// TIA Portal V20 export
// export: Created 2026-10-19T18:06:21.5238281Z, ExportSetting WithDefaults, DisplayName Totally Integrated Automation Portal, DisplayVersion V20 Update 6, DisplayName TIA Portal Openness, DisplayVersion V20 Update 6, DisplayName TIA Portal Version Control Interface, DisplayVersion V20 Update 6, DisplayName SINAMICS Startdrive Advanced, DisplayVersion V20 SP1, DisplayName SINAMICS Startdrive G130, G150, S120, S150, SINAMICS MV, G220, S200, S210, DisplayVersion V20 SP1, DisplayName SINAMICS Startdrive G110M, G120, G120C, G120D, G120P, G115D, DisplayVersion V20 SP1, DisplayName STEP 7 Professional, DisplayVersion V20 Update 6, DisplayName STEP 7 Safety, DisplayVersion V20 Update 2, DisplayName WinCC Basic/Comfort/Advanced, DisplayVersion V20 Update 6, DisplayName WinCC Unified, DisplayVersion V20 Update 6
FUNCTION_BLOCK "SAI_IND_CalFree"   // FB53, LAD
TITLE = CalFree Adjustment
{ S7_Optimized_Access := 'FALSE' }
VERSION : 0.1
// CalFree is a method of analog scale adjustment without using test weights. It takes the factory calibrated load cell Rated Output (mV/ Vexc.) and user defined scale capacity to build a linear loading curve.
// This method is usually applied to huge capacity scales in which calibration with test weights or other material is not feasible at all.
// stored: AutoNumber true, IsIECCheckEnabled false, SetENOAutomatically false, UDAEnableTagReadback false
   VAR_INPUT
      ID : HW_IO;   // The Profinet Device Hardware Identifier under device properties
   END_VAR
   VAR_OUTPUT
      Process : Bool;   // Adjustment is in process
      Done : Bool;   // Adjustment completed successfully
      Error : Bool;
   END_VAR
   VAR_IN_OUT
      RatedCapacity : Real;   // Scale Capacity
      Unit : SInt := 1;   // Decimal 0 - gram; 1 - KG; 2 - Lbs
      RatedOutput : Real;   // The averaged load cells' Rated Output in mV/V
      Start : Bool;   // Switch ON to start adjustment
   END_VAR
   VAR DB_SPECIFIC
      Activate : Bool;
      Status_RECORD : Int;
      CalFree_RECORD : Int;
      AdjustStep : SInt;
      Check01 : Bool;
      Check02 : Bool;
   END_VAR
   VAR
      WRREC_CalFree { S7_SetPoint := 'True'} : WRREC;
   END_VAR
   VAR DB_SPECIFIC
      Static01 : Bool;
   END_VAR
   VAR
      RDREC_Status { S7_SetPoint := 'True'} : RDREC;
   END_VAR
   VAR_TEMP   // added for the SCL form of the ladder/FBD networks
      _w1 : Bool;
      _w2 : Bool;
      _w3 : Bool;
      _w4 : Bool;
      _w5 : Bool;
      _w6 : Bool;
      _w7 : Bool;
      _w8 : Bool;
      _w9 : Bool;
      _w10 : Bool;
      _w11 : Bool;
   END_VAR
BEGIN

REGION Network 1: Start routine
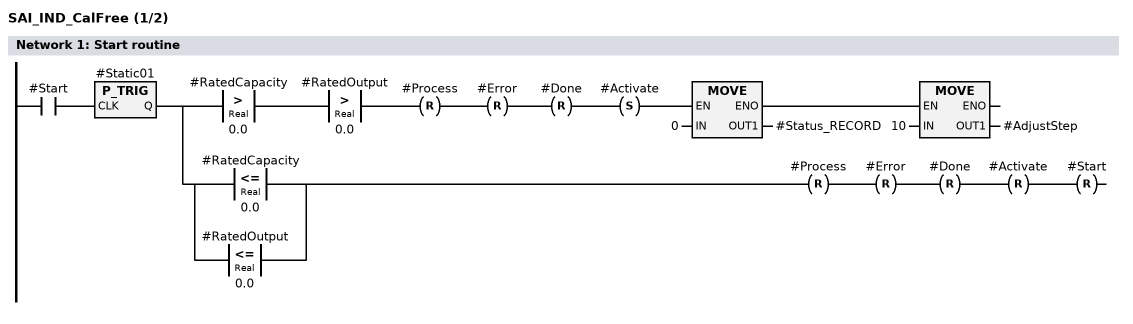
   RUNG wire#powerrail
      Contact( #Start )
      P_Trig( #Static01 )
      wire#w1
      { S7_Templates := "SrcType := Real" } GT_Contact(in1 := #RatedCapacity, in2 := 0.0)
      { S7_Templates := "SrcType := Real" } GT_Contact(in1 := #RatedOutput, in2 := 0.0)
      R_Coil( #Process )
      R_Coil( #Error )
      R_Coil( #Done )
      S_Coil( #Activate )
      Move(in := 0, out1 => #Status_RECORD)
      Move(in := 10, out1 => #AdjustStep)
   END_RUNG
   RUNG wire#w1
      { S7_Templates := "SrcType := Real" } LE_Contact(in1 := #RatedCapacity, in2 := 0.0)
      wire#w2
      R_Coil( #Process )
      R_Coil( #Error )
      R_Coil( #Done )
      R_Coil( #Activate )
      R_Coil( #Start )
   END_RUNG
   RUNG wire#w1
      { S7_Templates := "SrcType := Real" } LE_Contact(in1 := #RatedOutput, in2 := 0.0)
   END_RUNG wire#w2
   // the same network as SCL:
   #_w1 := #Start AND NOT #Static01;   // rising edge
   #Static01 := #Start;
   IF #_w1 AND (#RatedCapacity > 0.0) AND (#RatedOutput > 0.0) THEN
       #Process := FALSE;
       #Error := FALSE;
       #Done := FALSE;
       #Activate := TRUE;
       #Status_RECORD := 0;
       #AdjustStep := 10;
   END_IF;
   IF #_w1 AND ((#RatedCapacity <= 0.0) OR (#RatedOutput <= 0.0)) THEN
       #Process := FALSE;
       #Error := FALSE;
       #Done := FALSE;
       #Activate := FALSE;
       #Start := FALSE;
   END_IF;
END_REGION

REGION Network 2: Sequence
   // CalFree adjustment steps:
   // 
   // 1. Switch on Input bit Start
   // 
   // 2. Write in (a) Scale Capacity (Index 0x401A), (b) Scale unit (Index 0x401C, Decimal 0 - gram; Decimal 1 - KG; Decimal 2 - Pounds) and (c) Load Cells' averaged Rated Output (Index 0x401D, in mV/V)
   // 
   // 3. Start CalFree adjustment (Index 0x401A)
   // 
   // 4. Continuously read in adjustment status (Index 0x4007)
   // 
   // 5. Output bit Done will be turned ON after completion of the process
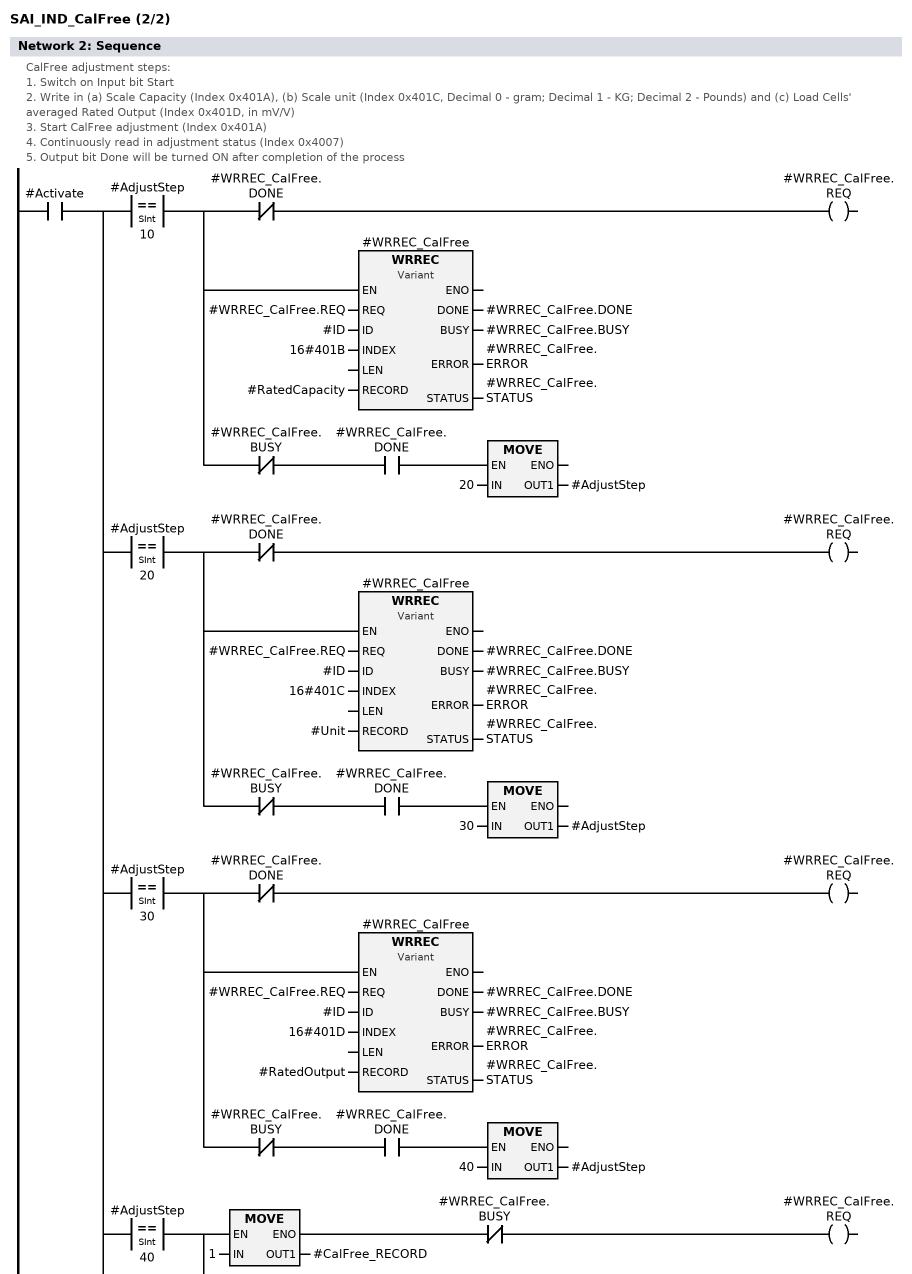
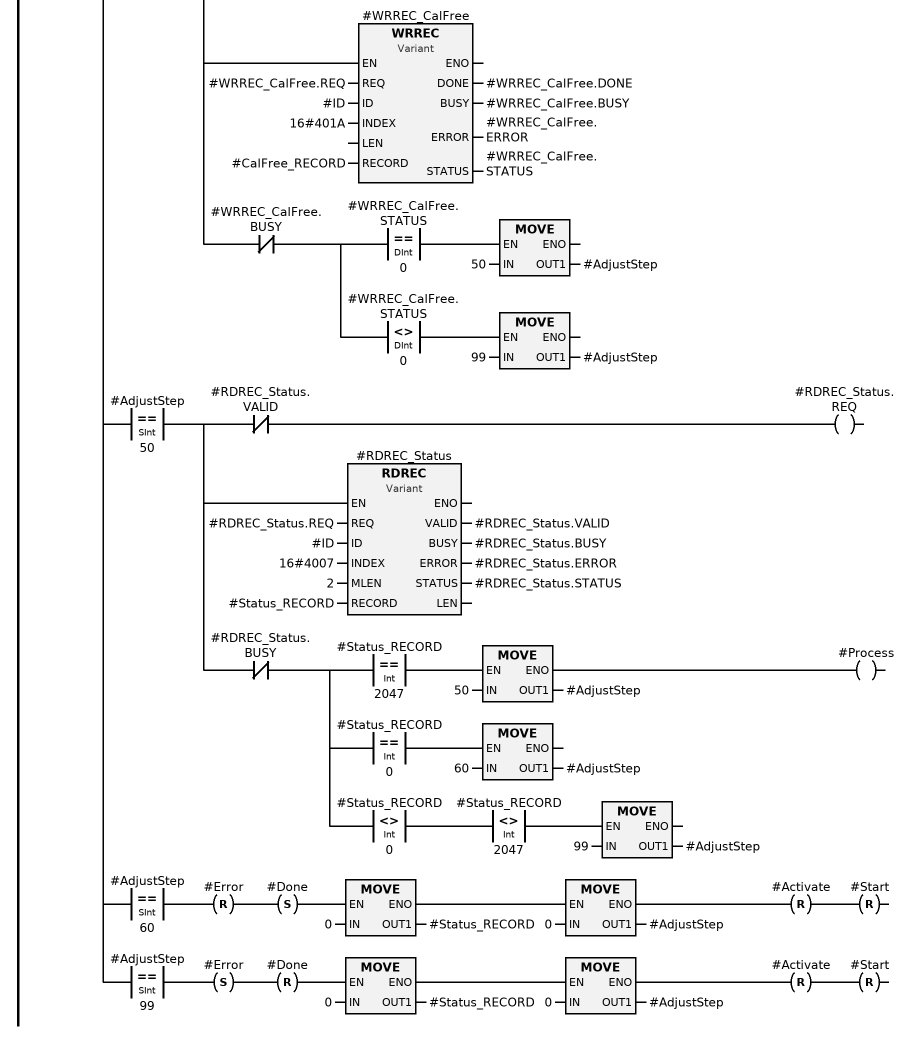
   RUNG wire#powerrail
      Contact( #Activate )
      wire#w1
      { S7_Templates := "SrcType := SInt" } EQ_Contact(in1 := #AdjustStep, in2 := 10)
      wire#w2
      I_Contact( #WRREC_CalFree.DONE )
      Coil( #WRREC_CalFree.REQ )
   END_RUNG
   RUNG wire#w2
      { S7_Templates := "[ptr_type := Variant, id_type := HW_IO, index_type := DInt, len_type := UInt]" } #WRREC_CalFree.WRREC(REQ := #WRREC_CalFree.REQ, ID := #ID, INDEX := 16#401B, LEN :=, RECORD := #RatedCapacity, DONE => #WRREC_CalFree.DONE, BUSY => #WRREC_CalFree.BUSY, ERROR => #WRREC_CalFree.ERROR, STATUS => #WRREC_CalFree.STATUS)
   END_RUNG
   RUNG wire#w2
      I_Contact( #WRREC_CalFree.BUSY )
      Contact( #WRREC_CalFree.DONE )
      Move(in := 20, out1 => #AdjustStep)
   END_RUNG
   RUNG wire#w1
      { S7_Templates := "SrcType := SInt" } EQ_Contact(in1 := #AdjustStep, in2 := 20)
      wire#w3
      I_Contact( #WRREC_CalFree.DONE )
      Coil( #WRREC_CalFree.REQ )
   END_RUNG
   RUNG wire#w3
      { S7_Templates := "[ptr_type := Variant, id_type := HW_IO, index_type := DInt, len_type := UInt]" } #WRREC_CalFree.WRREC(REQ := #WRREC_CalFree.REQ, ID := #ID, INDEX := 16#401C, LEN :=, RECORD := #Unit, DONE => #WRREC_CalFree.DONE, BUSY => #WRREC_CalFree.BUSY, ERROR => #WRREC_CalFree.ERROR, STATUS => #WRREC_CalFree.STATUS)
   END_RUNG
   RUNG wire#w3
      I_Contact( #WRREC_CalFree.BUSY )
      Contact( #WRREC_CalFree.DONE )
      Move(in := 30, out1 => #AdjustStep)
   END_RUNG
   RUNG wire#w1
      { S7_Templates := "SrcType := SInt" } EQ_Contact(in1 := #AdjustStep, in2 := 30)
      wire#w4
      I_Contact( #WRREC_CalFree.DONE )
      Coil( #WRREC_CalFree.REQ )
   END_RUNG
   RUNG wire#w4
      { S7_Templates := "[ptr_type := Variant, id_type := HW_IO, index_type := DInt, len_type := UInt]" } #WRREC_CalFree.WRREC(REQ := #WRREC_CalFree.REQ, ID := #ID, INDEX := 16#401D, LEN :=, RECORD := #RatedOutput, DONE => #WRREC_CalFree.DONE, BUSY => #WRREC_CalFree.BUSY, ERROR => #WRREC_CalFree.ERROR, STATUS => #WRREC_CalFree.STATUS)
   END_RUNG
   RUNG wire#w4
      I_Contact( #WRREC_CalFree.BUSY )
      Contact( #WRREC_CalFree.DONE )
      Move(in := 40, out1 => #AdjustStep)
   END_RUNG
   RUNG wire#w1
      { S7_Templates := "SrcType := SInt" } EQ_Contact(in1 := #AdjustStep, in2 := 40)
      wire#w5
      Move(in := 1, out1 => #CalFree_RECORD)
      I_Contact( #WRREC_CalFree.BUSY )
      Coil( #WRREC_CalFree.REQ )
   END_RUNG
   RUNG wire#w5
      { S7_Templates := "[ptr_type := Variant, id_type := HW_IO, index_type := DInt, len_type := UInt]" } #WRREC_CalFree.WRREC(REQ := #WRREC_CalFree.REQ, ID := #ID, INDEX := 16#401A, LEN :=, RECORD := #CalFree_RECORD, DONE => #WRREC_CalFree.DONE, BUSY => #WRREC_CalFree.BUSY, ERROR => #WRREC_CalFree.ERROR, STATUS => #WRREC_CalFree.STATUS)
   END_RUNG
   RUNG wire#w5
      I_Contact( #WRREC_CalFree.BUSY )
      wire#w6
      { S7_Templates := "SrcType := DInt" } EQ_Contact(in1 := #WRREC_CalFree.STATUS, in2 := 0)
      Move(in := 50, out1 => #AdjustStep)
   END_RUNG
   RUNG wire#w6
      { S7_Templates := "SrcType := DInt" } NE_Contact(in1 := #WRREC_CalFree.STATUS, in2 := 0)
      Move(in := 99, out1 => #AdjustStep)
   END_RUNG
   RUNG wire#w1
      { S7_Templates := "SrcType := SInt" } EQ_Contact(in1 := #AdjustStep, in2 := 50)
      wire#w7
      I_Contact( #RDREC_Status.VALID )
      Coil( #RDREC_Status.REQ )
   END_RUNG
   RUNG wire#w7
      { S7_Templates := "[ptr_type := Variant, id_type := HW_IO, index_type := DInt, len_type := UInt]" } #RDREC_Status.RDREC(REQ := #RDREC_Status.REQ, ID := #ID, INDEX := 16#4007, MLEN := 2, RECORD := #Status_RECORD, VALID => #RDREC_Status.VALID, BUSY => #RDREC_Status.BUSY, ERROR => #RDREC_Status.ERROR, STATUS => #RDREC_Status.STATUS, LEN =>)
   END_RUNG
   RUNG wire#w7
      I_Contact( #RDREC_Status.BUSY )
      wire#w8
      { S7_Templates := "SrcType := Int" } EQ_Contact(in1 := #Status_RECORD, in2 := 2047)
      Move(in := 50, out1 => #AdjustStep)
      Coil( #Process )
   END_RUNG
   RUNG wire#w8
      { S7_Templates := "SrcType := Int" } EQ_Contact(in1 := #Status_RECORD, in2 := 0)
      Move(in := 60, out1 => #AdjustStep)
   END_RUNG
   RUNG wire#w8
      { S7_Templates := "SrcType := Int" } NE_Contact(in1 := #Status_RECORD, in2 := 0)
      { S7_Templates := "SrcType := Int" } NE_Contact(in1 := #Status_RECORD, in2 := 2047)
      Move(in := 99, out1 => #AdjustStep)
   END_RUNG
   RUNG wire#w1
      { S7_Templates := "SrcType := SInt" } EQ_Contact(in1 := #AdjustStep, in2 := 60)
      R_Coil( #Error )
      S_Coil( #Done )
      Move(in := 0, out1 => #Status_RECORD)
      Move(in := 0, out1 => #AdjustStep)
      R_Coil( #Activate )
      R_Coil( #Start )
   END_RUNG
   RUNG wire#w1
      { S7_Templates := "SrcType := SInt" } EQ_Contact(in1 := #AdjustStep, in2 := 99)
      S_Coil( #Error )
      R_Coil( #Done )
      Move(in := 0, out1 => #Status_RECORD)
      Move(in := 0, out1 => #AdjustStep)
      R_Coil( #Activate )
      R_Coil( #Start )
   END_RUNG
   // the same network as SCL:
   #_w1 := #Activate AND (#AdjustStep = 10);
   #WRREC_CalFree.REQ := #_w1 AND NOT #WRREC_CalFree.DONE;
   IF #_w1 THEN
       #WRREC_CalFree(REQ := #WRREC_CalFree.REQ,   // WRREC
                      ID := #ID,
                      INDEX := 16#401B,
                      RECORD := #RatedCapacity,
                      DONE => #WRREC_CalFree.DONE,
                      BUSY => #WRREC_CalFree.BUSY,
                      ERROR => #WRREC_CalFree.ERROR,
                      STATUS => #WRREC_CalFree.STATUS);
   END_IF;
   IF #_w1 AND NOT #WRREC_CalFree.BUSY AND #WRREC_CalFree.DONE THEN #AdjustStep := 20; END_IF;
   #_w2 := #Activate AND (#AdjustStep = 20);
   #WRREC_CalFree.REQ := #_w2 AND NOT #WRREC_CalFree.DONE;
   IF #_w2 THEN
       #WRREC_CalFree(REQ := #WRREC_CalFree.REQ,   // WRREC
                      ID := #ID,
                      INDEX := 16#401C,
                      RECORD := #Unit,
                      DONE => #WRREC_CalFree.DONE,
                      BUSY => #WRREC_CalFree.BUSY,
                      ERROR => #WRREC_CalFree.ERROR,
                      STATUS => #WRREC_CalFree.STATUS);
   END_IF;
   IF #_w2 AND NOT #WRREC_CalFree.BUSY AND #WRREC_CalFree.DONE THEN #AdjustStep := 30; END_IF;
   #_w3 := #Activate AND (#AdjustStep = 30);
   #WRREC_CalFree.REQ := #_w3 AND NOT #WRREC_CalFree.DONE;
   IF #_w3 THEN
       #WRREC_CalFree(REQ := #WRREC_CalFree.REQ,   // WRREC
                      ID := #ID,
                      INDEX := 16#401D,
                      RECORD := #RatedOutput,
                      DONE => #WRREC_CalFree.DONE,
                      BUSY => #WRREC_CalFree.BUSY,
                      ERROR => #WRREC_CalFree.ERROR,
                      STATUS => #WRREC_CalFree.STATUS);
   END_IF;
   IF #_w3 AND NOT #WRREC_CalFree.BUSY AND #WRREC_CalFree.DONE THEN #AdjustStep := 40; END_IF;
   #_w4 := #Activate AND (#AdjustStep = 40);
   IF #_w4 THEN #CalFree_RECORD := 1; END_IF;
   #WRREC_CalFree.REQ := #_w4 AND NOT #WRREC_CalFree.BUSY;
   IF #_w4 THEN
       #WRREC_CalFree(REQ := #WRREC_CalFree.REQ,   // WRREC
                      ID := #ID,
                      INDEX := 16#401A,
                      RECORD := #CalFree_RECORD,
                      DONE => #WRREC_CalFree.DONE,
                      BUSY => #WRREC_CalFree.BUSY,
                      ERROR => #WRREC_CalFree.ERROR,
                      STATUS => #WRREC_CalFree.STATUS);
   END_IF;
   #_w5 := #_w4 AND NOT #WRREC_CalFree.BUSY;
   IF #_w5 AND (#WRREC_CalFree.STATUS = 0) THEN #AdjustStep := 50; END_IF;
   IF #_w5 AND (#WRREC_CalFree.STATUS <> 0) THEN #AdjustStep := 99; END_IF;
   #_w6 := #Activate AND (#AdjustStep = 50);
   #RDREC_Status.REQ := #_w6 AND NOT #RDREC_Status.VALID;
   IF #_w6 THEN
       #RDREC_Status(REQ := #RDREC_Status.REQ,   // RDREC
                     ID := #ID,
                     INDEX := 16#4007,
                     MLEN := 2,
                     RECORD := #Status_RECORD,
                     VALID => #RDREC_Status.VALID,
                     BUSY => #RDREC_Status.BUSY,
                     ERROR => #RDREC_Status.ERROR,
                     STATUS => #RDREC_Status.STATUS);
   END_IF;
   #_w7 := #_w6 AND NOT #RDREC_Status.BUSY;
   #_w8 := #_w7 AND (#Status_RECORD = 2047);
   IF #_w8 THEN #AdjustStep := 50; END_IF;
   #Process := #_w8;
   IF #_w7 AND (#Status_RECORD = 0) THEN #AdjustStep := 60; END_IF;
   IF #_w7 AND (#Status_RECORD <> 0) AND (#Status_RECORD <> 2047) THEN #AdjustStep := 99; END_IF;
   IF #Activate AND (#AdjustStep = 60) THEN
       #Error := FALSE;
       #Done := TRUE;
       #Status_RECORD := 0;
   END_IF;
   #_w9 := #Activate AND (#AdjustStep = 60);
   IF #_w9 THEN #AdjustStep := 0; END_IF;
   #_w10 := #Activate;
   IF #_w9 THEN
       #Activate := FALSE;
       #Start := FALSE;
   END_IF;
   IF #_w10 AND (#AdjustStep = 99) THEN
       #Error := TRUE;
       #Done := FALSE;
       #Status_RECORD := 0;
   END_IF;
   #_w11 := #_w10 AND (#AdjustStep = 99);
   IF #_w11 THEN
       #AdjustStep := 0;
       #Activate := FALSE;
       #Start := FALSE;
   END_IF;
END_REGION
END_FUNCTION_BLOCK
